(* IEC 61131-3 sources: Vigilimen/plant/plc-upload, 2 files *)

(* ---- conveyor_upload.st ---- *)
(*
    PLC-CONV-001 — control function for conveyor CONV-001
    Vigilimen · Sprint 3 · OpenPLC · Purdue Level 1, control zone

    This program sequences and protects the MACHINE. It does not protect
    people — SIS-CONV-001 does that, on a separate runtime, in a separate
    zone, with its own I/O, and this program has no path to it.

    Motor_Run below is a REQUEST. It is wired in series with the safety
    relay's contactor output, so:

        motor turns  =  safety contactor energised  AND  Motor_Run

    This program can stop the belt. It cannot start it against a trip.

    Reference model: plant/sim/interlock_model.py
    I/O contract:    plant/gateway/plc_io_map.py  (ADR-013), checked by FF-23
*)

PROGRAM PLC_CONV_001
VAR
    (* ── I/O contract with the gateway: plant/gateway/plc_io_map.py ────────
       FF-23 fails the build if this block and that table disagree.

       INPUTS. On a real plant these are physical inputs (%IX / %IW). Here
       the gateway plays the field over Modbus, and a Modbus master cannot
       write %IX or %IW, so the simulated field values live in %QX / %QW
       variables that this program only READS. It must never assign them:
       FF-23 checks that too. A simulation device, not a design to copy.
       Addresses 100+ are OpenPLC's slave range: coil = byte*8+bit, holding
       register = word number (ADR-013). *)
    Start_PB          AT %QX100.0 : BOOL;   (* start, local or SCADA          coil 800 *)
    Stop_PB           AT %QX100.1 : BOOL;   (* normal stop                    coil 801 *)
    Zero_Speed        AT %QX100.2 : BOOL;   (* TRUE when belt is stationary   coil 802 *)
    Upstream_Ready    AT %QX100.3 : BOOL;   (* crusher permissive             coil 803 *)
    Downstream_Ready  AT %QX100.4 : BOOL;   (* stockpile permissive           coil 804 *)
    Bearing_Temp_x10  AT %QW100   : UINT;   (* drive-end bearing, 0.1 degC    hreg 100 *)
    Motor_Current_x10 AT %QW101   : UINT;   (* amps x 10                      hreg 101 *)
    Belt_Speed_x100   AT %QW102   : UINT;   (* m/s x 100                      hreg 102 *)

    (* OUTPUTS. Written by this program, read by the gateway. *)
    Motor_Run         AT %QX101.0 : BOOL;   (* RUN REQUEST, in series with SIS coil 808 *)
    Alarm_Horn        AT %QX101.1 : BOOL;   (* pre-start warning              coil 809 *)
    Alarm_Word        AT %QW110   : WORD;   (* to SCADA                       hreg 110 *)
    Plc_State         AT %QW111   : UINT;   (* State below, for diagnostics   hreg 111 *)
    Plc_Map_Version   AT %QW112   : UINT;   (* signature: MAP_VERSION         hreg 112 *)
END_VAR

(* MatIEC (and the IEC grammar) takes a VAR block as ALL located or ALL plain.
   Mixing them in one block fails with 'invalid located variable declaration'
   on every plain line, then a cascade of ':=' errors (found by compiling in
   OpenPLC, 25 Oct). Located variables stay above; plain ones start here.
   FF-23 checks that no block mixes the two. *)
VAR
    (* Engineering values, decoded from the registers once per scan. *)
    Bearing_Temp    : REAL;    (* degC *)
    Motor_Current   : REAL;    (* amps *)
    Belt_Speed      : REAL;    (* m/s  *)

    State           : INT := 0;  (* 0 stopped 1 warning 2 starting 3 running 4 stopping 5 fault *)
    Warn_Timer      : TON;
    Start_Timer     : TON;
    Start_Edge      : R_TRIG;

    Permissives_OK  : BOOL;

    (* One BOOL per alarm bit. MatIEC does not accept bit access on a WORD
       (Alarm_Word.0 := ...), so the bits are kept separately and packed
       into Alarm_Word once per scan, at the end of the program.
       Bit 0 bearing, 1 current, 2 permissive, 3 start fail, 4 run stop. *)
    Alm_Bearing     : BOOL;
    Alm_Current     : BOOL;
    Alm_Permissive  : BOOL;
    Alm_StartFail   : BOOL;
    Alm_RunStop     : BOOL;
END_VAR

VAR CONSTANT
    BEARING_ALARM   : REAL := 85.0;
    BEARING_TRIP    : REAL := 95.0;
    OVERLOAD_TRIP   : REAL := 42.0;
    WARN_TIME       : TIME := T#10s;
    START_TIMEOUT   : TIME := T#15s;
    MAP_VERSION     : UINT := 1;   (* = plc_io_map.MAP_VERSION, FF-23 *)
END_VAR

(* ── Decode the registers ───────────────────────────────────────────── *)

Bearing_Temp  := UINT_TO_REAL(Bearing_Temp_x10) / 10.0;
Motor_Current := UINT_TO_REAL(Motor_Current_x10) / 10.0;
Belt_Speed    := UINT_TO_REAL(Belt_Speed_x100) / 100.0;

(* ── Permissives ────────────────────────────────────────────────────── *)

Permissives_OK := Upstream_Ready AND Downstream_Ready;

(* ── Machine protection ─────────────────────────────────────────────── *)

(* Alarms advise. Trips act. Both belong HERE and not in the safety
   function: they protect the conveyor, not a person, and a safety
   function loaded with machine protection trips more often for reasons
   operations do not respect. *)

Alm_Bearing    := Bearing_Temp >= BEARING_ALARM;
Alm_Current    := Motor_Current >= (OVERLOAD_TRIP * 0.9);
Alm_Permissive := NOT Permissives_OK;

IF Bearing_Temp >= BEARING_TRIP OR Motor_Current >= OVERLOAD_TRIP THEN
    State := 5;
END_IF;

(* ── Sequence ───────────────────────────────────────────────────────── *)

Start_Edge(CLK := Start_PB);

CASE State OF

0:  (* STOPPED *)
    Motor_Run  := FALSE;
    Alarm_Horn := FALSE;
    IF Start_Edge.Q AND Permissives_OK THEN
        State := 1;
    END_IF;

1:  (* PRE-START WARNING — the horn sounds before anything moves.
       A conveyor that starts silently is a conveyor someone is standing
       on. This delay is not politeness; it is the reason the belt is
       clear when it moves. *)
    Motor_Run  := FALSE;
    Alarm_Horn := TRUE;
    Warn_Timer(IN := TRUE, PT := WARN_TIME);
    IF Stop_PB THEN
        Warn_Timer(IN := FALSE);
        State := 0;
    ELSIF Warn_Timer.Q THEN
        Warn_Timer(IN := FALSE);
        State := 2;
    END_IF;

2:  (* STARTING — waiting for the belt to move *)
    Motor_Run  := TRUE;
    Alarm_Horn := FALSE;
    Start_Timer(IN := TRUE, PT := START_TIMEOUT);
    IF NOT Zero_Speed THEN
        Start_Timer(IN := FALSE);
        State := 3;
    ELSIF Start_Timer.Q THEN
        (* Commanded to run and did not move. Either the belt is stalled,
           or the SAFETY CONTACTOR IS OPEN — this program cannot tell the
           difference, and deliberately does not try. It stops asking. *)
        Start_Timer(IN := FALSE);
        Alm_StartFail := TRUE;
        State := 5;
    END_IF;

3:  (* RUNNING *)
    Motor_Run := TRUE;
    IF Stop_PB OR NOT Permissives_OK THEN
        State := 4;
    ELSIF Zero_Speed THEN
        (* Was running, now stationary, and nobody asked. Same reasoning
           as above: an unexplained stop is a fault, not a state to sit in *)
        Alm_RunStop   := TRUE;
        State := 5;
    END_IF;

4:  (* STOPPING *)
    Motor_Run := FALSE;
    IF Zero_Speed THEN
        State := 0;
    END_IF;

5:  (* FAULT — requires an operator acknowledgement, not a timer *)
    Motor_Run  := FALSE;
    Alarm_Horn := FALSE;
    IF Stop_PB AND Zero_Speed
       AND Bearing_Temp < BEARING_ALARM
       AND Motor_Current < 1.0
    THEN
        Alm_StartFail := FALSE;
        Alm_RunStop   := FALSE;
        State := 0;
    END_IF;

END_CASE;

Plc_State := INT_TO_UINT(State);
Plc_Map_Version := MAP_VERSION;

(* ── Pack the alarm bits for SCADA ──────────────────────────────────── *)

Alarm_Word := BOOL_TO_WORD(Alm_Bearing)
              OR SHL(BOOL_TO_WORD(Alm_Current), 1)
              OR SHL(BOOL_TO_WORD(Alm_Permissive), 2)
              OR SHL(BOOL_TO_WORD(Alm_StartFail), 3)
              OR SHL(BOOL_TO_WORD(Alm_RunStop), 4);

(*
    NOTE FOR THE 62443 ASSESSMENT AT S7

    Every input above arrives over Modbus TCP or S7comm. NEITHER PROTOCOL
    AUTHENTICATES ANYTHING. Anyone who can reach the port can write
    Start_PB, or Bearing_Temp, or Zero_Speed.

    That is not a defect in this program and cannot be fixed in it. It is
    why FR5 — restricted data flow — carries the weight it does in OT:
    the segmentation IS the authentication. See docs/architecture/
    protocol-register.md, and the write allow-list requirement that
    reaches the controller rather than the HMI.
*)

END_PROGRAM

(* ---------------------------------------------------------------------
   GENERATED by plant/plc-upload/build.py. Source: conveyor.st
   Only this block is added. Edit the source, then rebuild.
   --------------------------------------------------------------------- *)
CONFIGURATION Config0
  RESOURCE Res0 ON PLC
    TASK task0(INTERVAL := T#20ms, PRIORITY := 0);
    PROGRAM instance0 WITH task0 : PLC_CONV_001;
  END_RESOURCE
END_CONFIGURATION

(* ---- safety_upload.st ---- *)
(*
    SIS-CONV-001 — safety function for conveyor CONV-001
    Vigilimen · Sprint 3 · runs on OpenPLC, separate runtime, separate zone

    ─────────────────────────────────────────────────────────────────────
    THIS PROGRAM TAKES NO INPUT FROM THE CONTROL FUNCTION.

    There is no tag, no network path and no shared memory between this
    program and PLC-CONV-001. That is not a convention to be respected —
    it is enforced by the two running on separate runtimes, on separate
    zones, with separate I/O.

    Its output drops the motor contactor coil through a safety relay,
    wired in SERIES with the control PLC's motor output. The control
    function can stop the belt by dropping its own output. It cannot
    start the belt against this one, and it has no means of inhibiting,
    bypassing, delaying or acknowledging a trip.

    That asymmetry is the design. TRITON is why.
    ─────────────────────────────────────────────────────────────────────

    CONVENTION: TRUE = healthy / not demanded, on every input.
    De-energise to trip. A broken wire reads FALSE, which is a demand.
    Loss of power, loss of wire and a real demand all produce the same
    outcome — a trip mechanism that needs power to trip has a failure
    mode indistinguishable from normal operation.

    Reference model: plant/sim/interlock_model.py
    Verified by:     scripts/ff06_safety_independence.py  (13 cases)
    Settled by:      a witnessed test, and nothing else
*)

PROGRAM SIS_CONV_001
VAR_INPUT
    (* Dual-channel field devices. Two wires, two terminals, two reads. *)
    EStop_ChA       : BOOL;   (* %IX0.0  emergency stop, channel A     *)
    EStop_ChB       : BOOL;   (* %IX0.1  emergency stop, channel B     *)
    PullCord_ChA    : BOOL;   (* %IX0.2  belt pull-cord, channel A     *)
    PullCord_ChB    : BOOL;   (* %IX0.3  belt pull-cord, channel B     *)
    BeltDrift_OK    : BOOL;   (* %IX0.4  belt drift switch             *)
    Guard_Closed    : BOOL;   (* %IX0.5  guard position                *)
    Safety_Reset    : BOOL;   (* %IX0.6  MANUAL reset, at the panel    *)
END_VAR

VAR_OUTPUT
    Contactor_Coil  : BOOL;   (* %QX0.0  TRUE energises. Hardwired.    *)
    Trip_Latched    : BOOL;   (* %QX0.1  lamp at the panel             *)
    Device_Fault    : BOOL;   (* %QX0.2  discrepancy detected          *)
END_VAR

VAR
    (* Boots TRIPPED. A cold start is not a safe start: a controller that
       powers up permissive has decided the plant is safe without having
       looked at it. *)
    Tripped         : BOOL := TRUE;

    EStop_Demand    : BOOL;
    Cord_Demand     : BOOL;
    EStop_Discrep   : BOOL;
    Cord_Discrep    : BOOL;
    Discrep_Timer   : TON;
    Reset_Edge      : R_TRIG;
END_VAR

(* ── 1. Dual-channel evaluation ─────────────────────────────────────── *)

EStop_Demand  := NOT (EStop_ChA AND EStop_ChB);
Cord_Demand   := NOT (PullCord_ChA AND PullCord_ChB);

(* A discrepancy is a FAULT, not a vote.

   One channel healthy and one not means a broken wire or a welded
   contact. Either way the device can no longer be trusted to demand a
   stop WHEN IT IS NEEDED — which is a different and far worse failure
   than a spurious trip, because it is silent. *)

EStop_Discrep := EStop_ChA <> EStop_ChB;
Cord_Discrep  := PullCord_ChA <> PullCord_ChB;

Discrep_Timer(IN := (EStop_Discrep OR Cord_Discrep), PT := T#500ms);
Device_Fault  := Discrep_Timer.Q;

(* ── 2. Trip conditions ─────────────────────────────────────────────── *)

IF EStop_Demand
   OR Cord_Demand
   OR NOT BeltDrift_OK
   OR NOT Guard_Closed
   OR Device_Fault
THEN
    Tripped := TRUE;
END_IF;

(* ── 3. Reset ───────────────────────────────────────────────────────── *)

(* The trip LATCHES. Clearing the demand does not restart the belt:
   somebody pressed that stop and may now be standing at the machine.
   Reset is a rising edge at a physical panel button, not a level, and
   not a network write. *)

Reset_Edge(CLK := Safety_Reset);

IF Reset_Edge.Q
   AND NOT EStop_Demand
   AND NOT Cord_Demand
   AND BeltDrift_OK
   AND Guard_Closed
   AND NOT Device_Fault
THEN
    Tripped := FALSE;
END_IF;

(* ── 4. Output ──────────────────────────────────────────────────────── *)

Contactor_Coil := NOT Tripped;
Trip_Latched   := Tripped;

(*
    WHAT IS DELIBERATELY ABSENT, AND WHY

    No bearing temperature. No motor current. No vibration. No overload.

    Those are MACHINE protection and they live in PLC-CONV-001. Loading
    this program with them would add demands that have nothing to do with
    anyone's safety, and every added demand is another way for this
    function to trip spuriously — which is how a safety function ends up
    bypassed by people who need the plant to run.

    A safety function that trips for reasons operations do not respect
    will eventually be defeated, and then it protects nobody. Keeping it
    narrow is not minimalism. It is what keeps it trusted.

    No network input of any kind. No remote reset. No SCADA write.
    No "maintenance mode" bit. No bypass, timed or otherwise.
*)

END_PROGRAM

(* ---------------------------------------------------------------------
   GENERATED by plant/plc-upload/build.py. Source: safety.st
   Only this block is added. Edit the source, then rebuild.
   --------------------------------------------------------------------- *)
CONFIGURATION Config0
  RESOURCE Res0 ON PLC
    TASK task0(INTERVAL := T#20ms, PRIORITY := 0);
    PROGRAM instance0 WITH task0 : SIS_CONV_001;
  END_RESOURCE
END_CONFIGURATION
